Staubli VAL3: ListMove.pgx

public program ListMove(string x_sM)
  local bool l_bA
  local bool l_bB
  local bool l_bC
  local bool l_bEqual
  local joint l_jJoint
  local num l_nJogMode
  local jointRx l_jTargetPosUp
  local num l_nDir
  local point l_pTargetPosUp
  local point l_pCurrentPosUp
  local num l_nStep
  local bool l_bOut
  local trsf l_trA
  local trsf l_trB
  local point l_pA
  local pointRx l_pB
begin
  resetMotion()
  link(l_pCurrentPosUp,world)
  link(l_pTargetPosUp,world)
  //
  l_nJogMode=nJogMode
  $jogMode(0)
  wait($getJogmode()==0)
  delay(0.1)
  //
  //*******************************************************************************************
  switch x_sM
    case "pTeach1"
      call moveTarget(pTeach1,jTeach1)
    break
    //
    case "pTeach2"
      call moveTarget(pTeach2,jTeach2)
    break
    //
    case "pTeach3"
      call moveTarget(pTeach3,jTeach3)
    break
    //
    case "pTeach4"
      call moveTarget(pTeach4,jTeach4)
    break
    //
    case "pTeach5"
      call moveTarget(pTeach5,jTeach5)
    break
    //
    case "pTeach6"
      call moveTarget(pTeach6,jTeach6)
    break
    //
    case "pTeach7"
      call moveTarget(pTeach7,jTeach7)
    break
    //*******************************************************************************************
    case "pAdjustXY_2_1"
      call moveTarget(pAdjustXY_2_1,jAdjustXY_2_1)
    break
    //
    case "pAdjustXY_2_2"
      call moveTarget(pAdjustXY_2_2,jAdjustXY_2_2)
    break
    //
    case "pAdjustXY_3_1"
      call moveTarget(pAdjustXY_3_1,jAdjustXY_3_1)
    break
    //
    case "pAdjustXY_3_2"
      call moveTarget(pAdjustXY_3_2,jAdjustXY_3_2)
    break
    //
    case "pAdjustXY_3_3"
      call moveTarget(pAdjustXY_3_3,jAdjustXY_3_3)
    break
    //
    case "pAdjustZ_2_1"
      call moveTarget(pAdjustZ_2_1,jAdjustZ_2_1)
    break
    //
    case "pAdjustZ_2_2"
      call moveTarget(pAdjustZ_2_2,jAdjustZ_2_2)
    break
    //
    //*******************************************************************************************
    case "Align"
      call hmiAlert("Align","info")
      _pA.trsf={0,0,0,0,0,0}
      _pB.trsf={0,0,0,0,0,0}
      _pA=here(utCurrentTool.tValue,world)
      _pB=here(utCurrentTool.tValue,world)
      _pB.trsf=align(_pA.trsf,world.trsf)
      movel(_pB,utCurrentTool.tValue,mSpeed_C_blend)
      waitEndMove()
      call hmiAlert("CompleteAlign","info")
    break
    //
    case "GoBack_pAdjustXY_2_1"
      l_bOut=false
      l_nStep=0
      do
        switch l_nStep
          case 0
            if pAdjustXY_2_1.trsf!={0,0,0,0,0,0}
              l_nStep=1
            else
              l_nStep=99
            endIf
          break
          //
          case 1
            call CheckPosEqual(pAdjustXY_2_1,l_bEqual)
            if l_bEqual==true
              l_nStep=100
            else
              l_nStep=2
            endIf
          break
          //
          case 2
            call CheckPosEqual(pAdjustXY_2_2,l_bEqual)
            if l_bEqual==true
              l_nStep=3
            else
              l_nStep=4
            endIf
          break
          //
          case 3
            call hmiAlert("GoBack","info")
            movel(_pA,utCurrentTool.tValue,mSpeed_C_blend)
            movel(pAdjustXY_2_1,utCurrentTool.tValue,mSpeed_C_blend)
            waitEndMove()
            l_nStep=100
          break
          //
          case 4
            l_pCurrentPosUp=compose(here(utCurrentTool.tValue,world),world,{0,0,100*l_nDir,0,0,0})
            l_pTargetPosUp=appro(pAdjustXY_2_1,{0,0,-100,0,0,0})
            l_bA=pointToJoint(utCurrentTool.tValue,jAdjustXY_2_1,l_pTargetPosUp,l_jTargetPosUp)
            if l_bA==true
              call hmiAlert("GoBack","info")
              movel(l_pCurrentPosUp,utCurrentTool.tValue,mSpeed_J_blend)
              movej(l_jTargetPosUp,utCurrentTool.tValue,mSpeed_J_blend)
              movel(appro(pAdjustXY_2_1,{0,0,-20,0,0,0}),utCurrentTool.tValue,mSpeed_J_blend)
              movel(pAdjustXY_2_1,utCurrentTool.tValue,mSlow)
              waitEndMove()
              l_nStep=100
            else
              l_nStep=99
            endIf
          break
          //
          case 99
            call hmiAlert("CantGoBack","warning")
            l_bOut=true
          break
          //
          case 100
            call hmiAlert("CompleteGoBack","info")
            l_bOut=true
          break
        endSwitch
      until l_bOut
    break
    //
    case "Rz+180_pAdjustXY_2_1"
      l_bOut=false
      l_nStep=0
      do
        switch l_nStep
          case 0
            l_trA={0,0,0,0,0,90}
            l_trB={0,0,0,0,0,180}
            l_pA=appro(pAdjustXY_2_1,l_trA)
            l_pB=appro(pAdjustXY_2_1,l_trB)
            l_pA.config=cConfigSame
            l_pB.config=cConfigSame
            //
            call CheckPosEqual(l_pB,l_bEqual)
            if l_bEqual==true
              l_nStep=100
            else
              call CheckTraj(pAdjustXY_2_1,l_trA,l_pA,"Appro",l_bA)
              call CheckTraj(pAdjustXY_2_1,l_trB,l_pB,"Appro",l_bB)
              l_nStep=1
            endIf
          break
          //
          case 1
            //whether the target position is reachable
            if l_bA==true and l_bB==true
              l_nStep=2
            else
              l_nStep=99
            endIf
          break
          //
          case 2
            //Whether the robot is at the end position
            call CheckPosEqual(l_pB,l_bEqual)
            if !l_bEqual
              l_nStep=3
            else
              l_nStep=100
            endIf
          break
          //
          case 3
            call hmiAlert("Move","info")
            _pA=l_pA
            _pB=l_pB
            movel(_pA,utCurrentTool.tValue,mSpeed_C_blend)
            movel(_pB,utCurrentTool.tValue,mSpeed_C_blend)
            waitEndMove()
            l_nStep=100
          break
          //
          case 99
            call hmiAlert("CantMove1","warning")
            l_bOut=true
          break
          //
          case 100
            call hmiAlert("CompleteMove","info")
            l_bOut=true
          break
        endSwitch
      until l_bOut
    break
    //
    case "Rz-180_pAdjustXY_2_1"
      l_bOut=false
      l_nStep=0
      do
        switch l_nStep
          case 0
            l_trA={0,0,0,0,0,-90}
            l_trB={0,0,0,0,0,-180}
            l_pA=appro(pAdjustXY_2_1,l_trA)
            l_pB=appro(pAdjustXY_2_1,l_trB)
            l_pA.config=cConfigSame
            l_pB.config=cConfigSame
            //
            call CheckPosEqual(l_pB,l_bEqual)
            if l_bEqual==true
              l_nStep=100
            else
              call CheckTraj(pAdjustXY_2_1,l_trA,l_pA,"Appro",l_bA)
              call CheckTraj(pAdjustXY_2_1,l_trB,l_pB,"Appro",l_bB)
              l_nStep=1
            endIf
          break
          //
          case 1
            //whether the target position is reachable
            if l_bA==true and l_bB==true
              l_nStep=2
            else
              l_nStep=99
            endIf
          break
          //
          case 2
            //Whether the robot is at the end position
            call CheckPosEqual(l_pB,l_bEqual)
            if !l_bEqual
              l_nStep=3
            else
              l_nStep=100
            endIf
          break
          //
          case 3
            call hmiAlert("Move","info")
            _pA=l_pA
            _pB=l_pB
            movel(_pA,utCurrentTool.tValue,mSpeed_C_blend)
            movel(_pB,utCurrentTool.tValue,mSpeed_C_blend)
            waitEndMove()
            l_nStep=100
          break
          //
          case 99
            call hmiAlert("CantMove1","warning")
            l_bOut=true
          break
          //
          case 100
            call hmiAlert("CompleteMove","info")
            l_bOut=true
          break
        endSwitch
      until l_bOut
    break
    //
    case "GoBack_pAdjustXY_3_1"
      if pAdjustXY_3_1.trsf!={0,0,0,0,0,0}
        call CheckPosEqual(pAdjustXY_3_1,l_bEqual)
        if l_bEqual
          //At the starting positio
          call hmiAlert("CompleteGoBack","info")
        else
          //Not At the starting position
          call hmiAlert("GoBack","info")
          movel(pAdjustXY_3_1,utCurrentTool.tValue,mSpeed_C_blend)
          waitEndMove()
          call hmiAlert("CompleteGoBack","info")
        endIf
      else
        call hmiAlert("CantGoBack","warning")
      endIf
    break
    //
    case "Rz+60_pAdjustXY_3_1"
      l_bOut=false
      l_nStep=0
      do
        switch l_nStep
          case 0
            l_trA={0,0,0,0,0,60}
            _pA=appro(pAdjustXY_3_1,l_trA)
            _pA.config=cConfigSame
            //
            call CheckPosEqual(_pA,l_bEqual)
            if l_bEqual==true
              l_nStep=100
            else
              call CheckTraj(pAdjustXY_3_1,l_trA,_pA,"Appro",l_bA)
              l_nStep=1
            endIf
          break
          //
          case 1
            //whether the target position is reachable
            if l_bA==true
              l_nStep=2
            else
              l_nStep=99
            endIf
          break
          //
          case 2
            //Whether the robot is at the end position
            call CheckPosEqual(_pA,l_bEqual)
            if !l_bEqual
              l_nStep=3
            else
              l_nStep=100
            endIf
          break
          //
          case 3
            call hmiAlert("Move","info")
            movel(_pA,utCurrentTool.tValue,mSpeed_C_blend)
            waitEndMove()
            l_nStep=100
          break
          //
          case 99
            call hmiAlert("CantMove1","warning")
            l_bOut=true
          break
          //
          case 100
            call hmiAlert("CompleteMove","info")
            l_bOut=true
          break
        endSwitch
      until l_bOut
    break
    //
    case "Rz-60_pAdjustXY_3_1"
      l_bOut=false
      l_nStep=0
      do
        switch l_nStep
          case 0
            l_trA={0,0,0,0,0,-60}
            _pA=appro(pAdjustXY_3_1,l_trA)
            _pA.config=cConfigSame
            //
            call CheckPosEqual(_pA,l_bEqual)
            if l_bEqual==true
              l_nStep=100
            else
              call CheckTraj(pAdjustXY_3_1,l_trA,_pA,"Appro",l_bA)
              l_nStep=1
            endIf
          break
          //
          case 1
            //whether the target position is reachable
            if l_bA==true
              l_nStep=2
            else
              l_nStep=99
            endIf
          break
          //
          case 2
            //Whether the robot is at the end position
            call CheckPosEqual(_pA,l_bEqual)
            if !l_bEqual
              l_nStep=3
            else
              l_nStep=100
            endIf
          break
          //
          case 3
            call hmiAlert("Move","info")
            movel(_pA,utCurrentTool.tValue,mSpeed_C_blend)
            waitEndMove()
            l_nStep=100
          break
          //
          case 99
            call hmiAlert("CantMove1","warning")
            l_bOut=true
          break
          //
          case 100
            call hmiAlert("CompleteMove","info")
            l_bOut=true
          break
        endSwitch
      until l_bOut
    break
    //
    case "GoBack_pAdjustZ_2_1"
      if pAdjustZ_2_1.trsf!={0,0,0,0,0,0}
        call CheckPosEqual(pAdjustZ_2_1,l_bEqual)
        if l_bEqual
          //如果在起点
          call hmiAlert("CompleteGoBack","info")
        else
          //如果不在起点
          call hmiAlert("GoBack","info")
          movel(_pB,utCurrentTool.tValue,mSpeed_C_blend)
          movel(pAdjustZ_2_1,utCurrentTool.tValue,mSlow)
          waitEndMove()
          call hmiAlert("CompleteGoBack","info")
        endIf
      else
        call hmiAlert("CantGoBack","warning")
      endIf
    break
    //
    case "Rx+60_pAdjustZ_2_1"
      l_bOut=false
      l_nStep=0
      do
        switch l_nStep
          case 0
            l_trA={0,0,0,60,0,0}
            l_pA=compose(pAdjustZ_2_1,world,l_trA)
            l_pA.trsf.x=pAdjustZ_2_1.trsf.x
            l_pA.trsf.y=pAdjustZ_2_1.trsf.y
            l_pA.trsf.z=pAdjustZ_2_1.trsf.z
            l_pB=appro(pAdjustZ_2_1,{0,0,-10,0,0,0})
            l_pA.config=cConfigSame
            l_pB.config=cConfigSame
            //
            call CheckPosEqual(l_pA,l_bEqual)
            if l_bEqual==true
              l_nStep=100
            else
              call CheckTraj(pAdjustZ_2_1,l_trB,l_pB,"Appro",l_bA)
              call CheckTraj(l_pB,l_trA,l_pA,"Compose",l_bB)
              l_nStep=1
            endIf
          break
          //
          case 1
            //whether the target position is reachable
            if l_bA==true and l_bB==true
              l_nStep=2
            else
              l_nStep=99
            endIf
          break
          //
          case 2
            //Whether the robot is at the end position
            call CheckPosEqual(l_pB,l_bEqual)
            if !l_bEqual
              l_nStep=3
            else
              l_nStep=100
            endIf
          break
          //
          case 3
            call hmiAlert("Move","info")
            _pA=l_pA
            _pB=l_pB
            movel(_pB,utCurrentTool.tValue,mSpeed_C_blend)
            movel(_pA,utCurrentTool.tValue,mSpeed_C_blend)
            waitEndMove()
            l_nStep=100
          break
          //
          case 99
            call hmiAlert("CantMove1","warning")
            l_bOut=true
          break
          //
          case 100
            call hmiAlert("CompleteMove","info")
            l_bOut=true
          break
        endSwitch
      until l_bOut
    break
    //
    case "Ry+60_pAdjustZ_2_1"
      l_bOut=false
      l_nStep=0
      do
        switch l_nStep
          case 0
            l_trA={0,0,0,0,60,0}
            l_pA=compose(pAdjustZ_2_1,world,l_trA)
            l_pA.trsf.x=pAdjustZ_2_1.trsf.x
            l_pA.trsf.y=pAdjustZ_2_1.trsf.y
            l_pA.trsf.z=pAdjustZ_2_1.trsf.z
            l_pB=appro(pAdjustZ_2_1,{0,0,-10,0,0,0})
            l_pA.config=cConfigSame
            l_pB.config=cConfigSame
            //
            call CheckPosEqual(l_pA,l_bEqual)
            if l_bEqual==true
              l_nStep=100
            else
              call CheckTraj(pAdjustZ_2_1,l_trB,l_pB,"Appro",l_bA)
              call CheckTraj(l_pB,l_trA,l_pA,"Compose",l_bB)
              l_nStep=1
            endIf
          break
          //
          case 1
            //whether the target position is reachable
            if l_bA==true and l_bB==true
              l_nStep=2
            else
              l_nStep=99
            endIf
          break
          //
          case 2
            //Whether the robot is at the end position
            call CheckPosEqual(l_pB,l_bEqual)
            if !l_bEqual
              l_nStep=3
            else
              l_nStep=100
            endIf
          break
          //
          case 3
            call hmiAlert("Move","info")
            _pA=l_pA
            _pB=l_pB
            movel(_pB,utCurrentTool.tValue,mSpeed_C_blend)
            movel(_pA,utCurrentTool.tValue,mSpeed_C_blend)
            waitEndMove()
            l_nStep=100
          break
          //
          case 99
            call hmiAlert("CantMove1","warning")
            l_bOut=true
          break
          //
          case 100
            call hmiAlert("CompleteMove","info")
            l_bOut=true
          break
        endSwitch
      until l_bOut
    break
  endSwitch
  $jogMode(l_nJogMode)
end
